// TIA Portal V20 export
// export: Created 2026-10-06T00:00:00
ScreenTemplate "Base"  1280x800, Number=1
  ScreenLayer 
    Rectangle "Header" at 0,100 size 40x40
